Yaskawa INFORM job: NAMEPRO.JBI

/JOB
//NAME NAMEPRO
//POS
///NPOS 6,0,0,0,0,0
///TOOL 9
///POSTYPE PULSE
///PULSE
C00000=0,0,0,0,0,0
C00001=0,0,0,0,0,0
C00002=0,0,0,0,0,0
C00003=0,0,0,0,0,0
C00004=0,0,0,0,0,0
C00005=0,0,0,0,0,0
//INST
<volatile>
///COMM Generated using RoboDK
///ATTR SC,RW
///GROUP1 RB1
NOP
'Program generated by RoboDK v
'6.0.7 for Yaskawa Motoman EPL
'160 on XX/XX/XXXX 18:00:00
'Using nominal kinematics.
'Using Frame S (targets wrt ba
'se):
'1234.6,-98.8,50.5,0.0,0.0,30.
'0
'Tool Tool S should be close t
'o:
'10.0,20.0,150.0,0.0,0.0,0.0
MOVJ C00000 VJ=50.00
MOVL C00001 V=100.0
MOVC C00002 V=100.0
MOVC C00003 V=100.0
MOVC C00004 V=100.0
MOVJ C00005 VJ=50.00
END
